// TIA Portal V21 export
// export: Created 2026-08-21T20:18:56.7717211Z, ExportSetting None, DisplayName Totally Integrated Automation Portal, DisplayVersion V21, DisplayName STEP 7 Professional, DisplayVersion V21, DisplayName STEP 7 Safety, DisplayVersion V21, DisplayName Tech WebApplication, DisplayVersion V21, DisplayName WinCC Basic/Comfort/Advanced, DisplayVersion V21, DisplayName WinCC Professional, DisplayVersion V21, DisplayName WinCC Unified, DisplayVersion V21
TYPE "UDT_Service_ParameterDefinition"
   STRUCT
      indexMTP : Int;   // Index of parameter / MTP Index of parameter
      indexIO : Int;   // Index of parameter / IO Index of parameter
      "type" : Int;   // Type of parameter
      controlModule : Byte := 16#FF;   // Number of control module used with parameter
   END_STRUCT;
END_TYPE
